% RSLogix 500 project Automatic Motor Stop Timer_BAK006.RSS, saved by version 8.30.00.16 %
PROJECT "PLCLAB"    % processor: Bul.1763 MicroLogix 1100 Series B %

PROGRAM FILES
  LAD 2 "MAIN"  5 rungs
  LAD 3 "DIGITAL IO"  4 rungs
  LAD 4 "ANALOG IO"  1 rungs
  LAD 5 "ALARMS"  1 rungs
  LAD 6 "CONTROLS"  4 rungs

DATA FILES
  O0 OUTPUT  5 elements
  I1 INPUT  7 elements
  S2 STATUS  66 elements
  B3 BINARY  1 elements
  T4 TIMER  1 elements
  C5 COUNTER  1 elements
  R6 CONTROL  1 elements
  N7 INTEGER  1 elements
  F8 FLOAT  1 elements

LADDER 2 "MAIN"
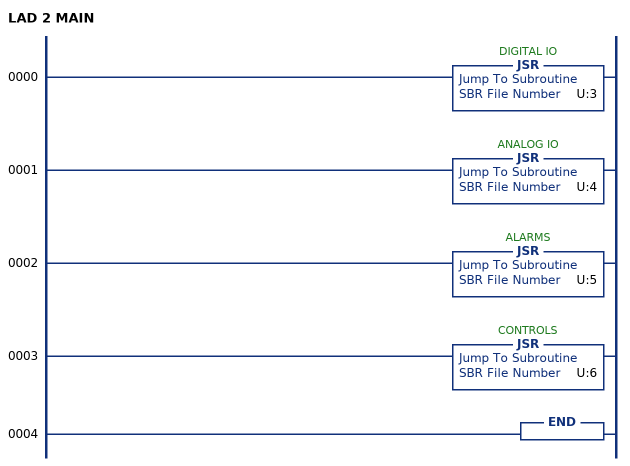
% Rung: 0 %
SOR JSR U:3 EOR
%   U:3  "DIGITAL IO" %
% Rung: 1 %
SOR JSR U:4 EOR
%   U:4  "ANALOG IO" %
% Rung: 2 %
SOR JSR U:5 EOR
%   U:5  "ALARMS" %
% Rung: 3 %
SOR JSR U:6 EOR
%   U:6  "CONTROLS" %
% Rung: 4 %
SOR END EOR

LADDER 3 "DIGITAL IO"
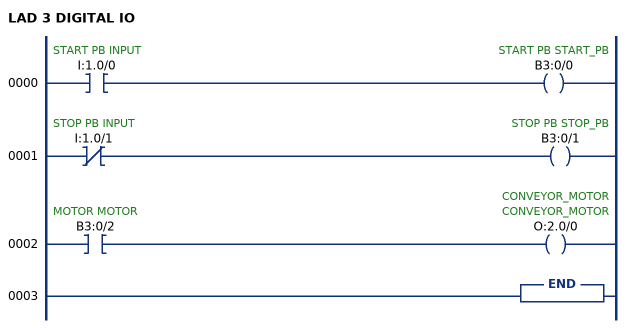
% Rung: 0 %
SOR XIC I:1.0/0 OTE B3:0/0 EOR
%   I:1.0/0  "START PB INPUT" %
%   B3:0/0  START_PB  "START PB" %
% Rung: 1 %
SOR XIO I:1.0/1 OTE B3:0/1 EOR
%   I:1.0/1  "STOP PB INPUT" %
%   B3:0/1  STOP_PB  "STOP PB" %
% Rung: 2 %
SOR XIC B3:0/2 OTE O:2.0/0 EOR
%   B3:0/2  MOTOR  "MOTOR" %
%   O:2.0/0  CONVEYOR_MOTOR  "CONVEYOR_MOTOR" %
% Rung: 3 %
SOR END EOR

LADDER 6 "CONTROLS"
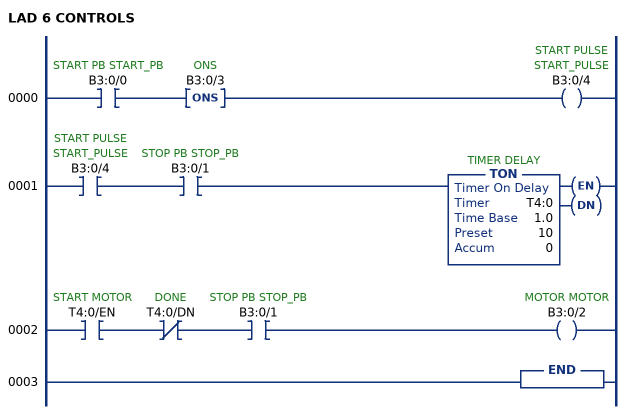
% Rung: 0 %
SOR XIC B3:0/0 ONS B3:0/3 OTE B3:0/4 EOR
%   B3:0/0  START_PB  "START PB" %
%   B3:0/3  "ONS" %
%   B3:0/4  START_PULSE  "START PULSE" %
% Rung: 1 %
SOR XIC B3:0/4 XIC B3:0/1 TON T4:0 1.0 10 0 EOR
%   B3:0/4  START_PULSE  "START PULSE" %
%   B3:0/1  STOP_PB  "STOP PB" %
%   T4:0  "TIMER DELAY" %
% Rung: 2 %
SOR XIC T4:0/EN XIO T4:0/DN XIC B3:0/1 OTE B3:0/2 EOR
%   T4:0/EN  "START MOTOR" %
%   T4:0/DN  "DONE" %
%   B3:0/1  STOP_PB  "STOP PB" %
%   B3:0/2  MOTOR  "MOTOR" %
% Rung: 3 %
SOR END EOR

DATA TABLE (non-zero values as saved)
DATA T4
% .PRE .ACC %
% T4:0 % 10 0
